Fanuc KAREL source: KB00106.KL

PROGRAM KB00106
%NOLOCKGROUP
%ENVIRONMENT PBQMGR
VAR
  P1: QUEUE_TYPE
BEGIN
  INIT_QUEUE(P1)
END KB00106
